ORGANIZATION_BLOCK FC 1
BEGIN
END_ORGANIZATION_BLOCK
